TYPE "ST_DeclarationParCmd"
VERSION : 0.1
   STRUCT
      Value : DInt;
   END_STRUCT;

END_TYPE

